            num nMoveType = 4
            num nPercentage
            num nSigValue = 1
        pointRx pPointRx[2]
        string sID
      [2]
        bool bMarked
        jointRx jJointRx = {j1=-87.551314, j2=145.129335, j3=-83.0857287, j4=182.11845, j5=63.691242, j6=-64.966659}
        pointRx pInter
        paraItem pParaItem
          [0]
            bool bSafePoint
            ifItem iIfItem
              [0]
                bool bANDOR[2]
                num nSigIndex[3]
                num nSigType[3]
                num nValue[3]
            mdesc mMdesc
            num nActionIndex = 42
            num nDelay
            num nMoveType = 1
            num nPercentage
            num nSigValue = 1
        pointRx pPointRx[2] = {x=61.349727, y=-652.129552, z=350.0734551, rx=-1.549449, ry=-1.96692, rz=28.421736, shoulder=lefty, elbow=enegative, wrist=wpositive}
        string sID
      [3]
        bool bMarked
        jointRx jJointRx = {j1=-47.00566362, j2=123.661152, j3=-79.978164, j4=176.739672, j5=50.379836, j6=-102.275032}
        pointRx pInter
        paraItem pParaItem
          [0]
            bool bSafePoint
            ifItem iIfItem
              [0]
                bool bANDOR[2]
                num nSigIndex[3]
                num nSigType[3]
                num nValue[3]
            mdesc mMdesc
            num nActionIndex = 42
            num nDelay
            num nMoveType = 1
            num nPercentage
            num nSigValue = 1
        pointRx pPointRx[2] = {x=488.627273, y=-418.649607, z=567.937104, rx=-6.582637, ry=-2.686226, rz=28.338446, shoulder=lefty, elbow=enegative, wrist=wpositive}
        string sID
      [4]
        bool bMarked
        jointRx jJointRx = {j1=-49.0942088, j2=121.00459063, j3=-74.169176, j4=177.183335, j5=53.609232, j6=-100.608132}
        pointRx pInter
        paraItem pParaItem
          [0]
            bool bSafePoint
            ifItem iIfItem
              [0]
                bool bANDOR[2]
                num nSigIndex[3]
                num nSigType[3]
                num nValue[3]
            mdesc mMdesc
            num nActionIndex = 42
            num nDelay
            num nMoveType = 1
            num nPercentage
            num nSigValue = 1
        pointRx pPointRx[2] = {x=488.602234, y=-457.380545, z=567.975681, rx=-6.584679, ry=-2.688341, rz=28.337484, shoulder=lefty, elbow=enegative, wrist=wpositive}
        string sID
      [5]
        bool bMarked
        jointRx jJointRx = {j1=-49.663191, j2=124.62488, j3=-82.121571, j4=177.0975297, j5=49.304971, j6=-99.821288}
        pointRx pInter
        paraItem pParaItem
          [0]
            bool bSafePoint
            ifItem iIfItem
              [0]
                bool bANDOR[2]
                num nSigIndex[3]
                num nSigType[3]
                num nValue[3]
            mdesc mMdesc
            num nActionIndex = 42
            num nDelay
            num nMoveType = 1
            num nPercentage
            num nSigValue = 1
        pointRx pPointRx[2] = {x=459.245528, y=-433.916408, z=567.993278, rx=-6.586651, ry=-2.689923, rz=28.337206, shoulder=lefty, elbow=enegative, wrist=wpositive}
        string sID
      [6]
        bool bMarked
        jointRx jJointRx = {j1=-51.089262, j2=127.485832, j3=-88.52739, j4=177.166583, j5=45.811078, j6=-98.322007}
        pointRx pInter
        paraItem pParaItem
          [0]
            bool bSafePoint
            ifItem iIfItem
              [0]
                bool bANDOR[2]
                num nSigIndex[3]
                num nSigType[3]
                num nValue[3]
            mdesc mMdesc
            num nActionIndex = 42
            num nDelay
            num nMoveType = 1
            num nPercentage
            num nSigValue = 1
        pointRx pPointRx[2] = {x=426.511567, y=-420.559077, z=567.993292, rx=-6.586458, ry=-2.69014, rz=28.337108, shoulder=lefty, elbow=enegative, wrist=wpositive}
        string sID
      [7]
        bool bMarked
        jointRx jJointRx = {j1=-53.0755743, j2=125.0272638, j3=-83.0148913, j4=177.619487, j5=48.919255, j6=-96.759929}
        pointRx pInter
        paraItem pParaItem
          [0]
            bool bSafePoint
            ifItem iIfItem
              [0]
                bool bANDOR[2]
                num nSigIndex[3]
                num nSigType[3]
                num nValue[3]
            mdesc mMdesc
            num nActionIndex = 42
            num nDelay
            num nMoveType = 1
            num nPercentage
            num nSigValue = 1
        pointRx pPointRx[2] = {x=426.51149, y=-458.270304, z=567.99328, rx=-6.585479, ry=-2.689619, rz=28.337033, shoulder=lefty, elbow=enegative, wrist=wpositive}
        string sID
      [8]
        bool bMarked
        jointRx jJointRx = {j1=-52.426636, j2=130.387774, j3=-95.172697, j4=177.208528, j5=42.11144, j6=-96.897847}
        pointRx pInter
        paraItem pParaItem
          [0]
            bool bSafePoint
            ifItem iIfItem
              [0]
                bool bANDOR[2]
                num nSigIndex[3]
                num nSigType[3]
                num nValue[3]
            mdesc mMdesc
            num nActionIndex = 42
            num nDelay
            num nMoveType = 1
            num nPercentage
            num nSigValue = 1
        pointRx pPointRx[2] = {x=393.481918, y=-402.66269, z=567.993281, rx=-6.585883, ry=-2.690348, rz=28.336908, shoulder=lefty, elbow=enegative, wrist=wpositive}
        string sID
      [9]
        bool bMarked
        jointRx jJointRx = {j1=-58.974439, j2=129.367388, j3=-92.816655, j4=178.435502, j5=43.592863, j6=-91.334255}
        pointRx pInter
        paraItem pParaItem
          [0]
            bool bSafePoint
            ifItem iIfItem
              [0]
                bool bANDOR[2]
                num nSigIndex[3]
                num nSigType[3]
                num nValue[3]
            mdesc mMdesc
            num nActionIndex = 42
            num nDelay
            num nMoveType = 1
            num nPercentage
            num nSigValue = 1
        pointRx pPointRx[2] = {x=344.945517, y=-458.235382, z=567.993294, rx=-6.587043, ry=-2.691097, rz=28.336907, shoulder=lefty, elbow=enegative, wrist=wpositive}
        string sID
      [10]
        bool bMarked
        jointRx jJointRx = {j1=-57.192018, j2=131.638959, j3=-98.096273, j4=178.00498558, j5=40.554749, j6=-92.720675}
        pointRx pInter
        paraItem pParaItem
          [0]
            bool bSafePoint
            ifItem iIfItem
              [0]
                bool bANDOR[2]
                num nSigIndex[3]
                num nSigType[3]
                num nValue[3]
            mdesc mMdesc
            num nActionIndex = 42
            num nDelay
            num nMoveType = 1
            num nPercentage
            num nSigValue = 1
        pointRx pPointRx[2] = {x=344.980685, y=-421.973821, z=567.993293, rx=-6.587471, ry=-2.690641, rz=28.337121, shoulder=lefty, elbow=enegative, wrist=wpositive}
        string sID
      [11]
        bool bMarked
        jointRx jJointRx = {j1=-60.376179, j2=132.512186, j3=-100.160991, j4=178.57184, j5=39.414626, j6=-89.972735}
        pointRx pInter
        paraItem pParaItem
          [0]
            bool bSafePoint
            ifItem iIfItem
              [0]
                bool bANDOR[2]
                num nSigIndex[3]
                num nSigType[3]
                num nValue[3]
            mdesc mMdesc
            num nActionIndex = 42
            num nDelay
            num nMoveType = 1
            num nPercentage
            num nSigValue = 1
        pointRx pPointRx[2] = {x=311.978155, y=-431.490165, z=567.993281, rx=-6.586244, ry=-2.690739, rz=28.336894, shoulder=lefty, elbow=enegative, wrist=wpositive}
        string sID
      [12]
        bool bMarked
        jointRx jJointRx = {j1=-65.107588, j2=132.458168, j3=-100.0326711, j4=179.493071, j5=39.531997, j6=-85.98983}
        pointRx pInter
        paraItem pParaItem
          [0]
            bool bSafePoint
            ifItem iIfItem
              [0]
                bool bANDOR[2]
                num nSigIndex[3]
                num nSigType[3]
                num nValue[3]
            mdesc mMdesc
            num nActionIndex = 42
            num nDelay
            num nMoveType = 1
            num nPercentage
            num nSigValue = 1
        pointRx pPointRx[2] = {x=270.822712, y=-458.161765, z=567.993281, rx=-6.586253, ry=-2.691371, rz=28.336679, shoulder=lefty, elbow=enegative, wrist=wpositive}
        string sID
      [13]
        bool bMarked
        jointRx jJointRx = {j1=-63.595033, j2=134.613161, j3=-105.229763, j4=179.141794, j5=36.481622, j6=-87.191501}
        pointRx pInter
        paraItem pParaItem
          [0]
            bool bSafePoint
            ifItem iIfItem
              [0]
                bool bANDOR[2]
                num nSigIndex[3]
                num nSigType[3]
                num nValue[3]
            mdesc mMdesc
            num nActionIndex = 42
            num nDelay
            num nMoveType = 1
            num nPercentage
            num nSigValue = 1
        pointRx pPointRx[2] = {x=270.822707, y=-423.00547317, z=567.99328, rx=-6.587117, ry=-2.691103, rz=28.336883, shoulder=lefty, elbow=enegative, wrist=wpositive}
        string sID
      [14]
        bool bMarked
        jointRx jJointRx = {j1=-65.403022, j2=136.841875, j3=-110.804443, j4=179.476622, j5=33.145897, j6=-85.649351}
        pointRx pInter
        paraItem pParaItem
          [0]
            bool bSafePoint
            ifItem iIfItem
              [0]
                bool bANDOR[2]
                num nSigIndex[3]
                num nSigType[3]
                num nValue[3]
            mdesc mMdesc
            num nActionIndex = 42
            num nDelay
            num nMoveType = 1
            num nPercentage
            num nSigValue = 1
        pointRx pPointRx[2] = {x=241.448098, y=-401.317138, z=567.99328, rx=-6.586652, ry=-2.691495, rz=28.336732, shoulder=lefty, elbow=enegative, wrist=wpositive}
        string sID
      [15]
        bool bMarked
        jointRx jJointRx = {j1=-71.552923, j2=137.207285, j3=-111.742738, j4=180.882707, j5=32.563572, j6=-80.728949}
        pointRx pInter
        paraItem pParaItem
          [0]
            bool bSafePoint
            ifItem iIfItem
              [0]
                bool bANDOR[2]
                num nSigIndex[3]
                num nSigType[3]
                num nValue[3]
            mdesc mMdesc
            num nActionIndex = 42
            num nDelay
            num nMoveType = 1
            num nPercentage
            num nSigValue = 1
        pointRx pPointRx[2] = {x=188.956768, y=-421.559208, z=567.993271, rx=-6.585305, ry=-2.691208, rz=28.336687, shoulder=lefty, elbow=enegative, wrist=wpositive}
        string sID
      [16]
        bool bMarked
        jointRx jJointRx = {j1=-72.731137, j2=135.0432437, j3=-106.287062, j4=181.0587207, j5=35.845376, j6=-79.673802}
        pointRx pInter
        paraItem pParaItem
          [0]
            bool bSafePoint
            ifItem iIfItem
              [0]
                bool bANDOR[2]
                num nSigIndex[3]
                num nSigType[3]
                num nValue[3]
            mdesc mMdesc
            num nActionIndex = 42
            num nDelay
            num nMoveType = 1
            num nPercentage
            num nSigValue = 1
        pointRx pPointRx[2] = {x=188.956768, y=-457.62638, z=567.99327, rx=-6.585271, ry=-2.690608, rz=28.336851, shoulder=lefty, elbow=enegative, wrist=wpositive}
        string sID
      [17]
        bool bMarked
        jointRx jJointRx = {j1=-75.0748224, j2=137.195165, j3=-111.715211, j4=181.688824, j5=32.546968, j6=-77.913471}
        pointRx pInter
        paraItem pParaItem
          [0]
            bool bSafePoint
            ifItem iIfItem
              [0]
                bool bANDOR[2]
                num nSigIndex[3]
                num nSigType[3]
                num nValue[3]
            mdesc mMdesc
            num nActionIndex = 42
            num nDelay
            num nMoveType = 1
            num nPercentage
            num nSigValue = 1
        pointRx pPointRx[2] = {x=159.184051, y=-433.850025, z=568.00311248, rx=-6.587391, ry=-2.691219, rz=28.336525, shoulder=lefty, elbow=enegative, wrist=wpositive}
        string sID
      [18]
        bool bMarked
        jointRx jJointRx = {j1=-79.693745, j2=136.402957, j3=-109.689565, j4=182.654161, j5=33.70043, j6=-74.112995}
        pointRx pInter
        paraItem pParaItem
          [0]
            bool bSafePoint
            ifItem iIfItem
              [0]
                bool bANDOR[2]
                num nSigIndex[3]
                num nSigType[3]
                num nValue[3]
            mdesc mMdesc
            num nActionIndex = 42
            num nDelay
            num nMoveType = 1
            num nPercentage
            num nSigValue = 1
        pointRx pPointRx[2] = {x=121.279103, y=-459.277382, z=568.00309762, rx=-6.585667, ry=-2.690876, rz=28.336551, shoulder=lefty, elbow=enegative, wrist=wpositive}
        string sID
      [19]
        bool bMarked
        jointRx jJointRx = {j1=-78.970374, j2=138.503231, j3=-115.146628, j4=182.739047, j5=30.363076, j6=-74.986334}
        pointRx pInter
        paraItem pParaItem
          [0]
            bool bSafePoint
            ifItem iIfItem
              [0]
                bool bANDOR[2]
                num nSigIndex[3]
                num nSigType[3]
                num nValue[3]
            mdesc mMdesc
            num nActionIndex = 42
            num nDelay
            num nMoveType = 1
            num nPercentage
            num nSigValue = 1
        pointRx pPointRx[2] = {x=121.279109, y=-423.991398, z=568.0031016, rx=-6.587075, ry=-2.690729, rz=28.336634, shoulder=lefty, elbow=enegative, wrist=wpositive}
        string sID
      [20]
        bool bMarked
        jointRx jJointRx = {j1=-82.18311, j2=140.325944, j3=-120.168865, j4=183.894102, j5=27.100815, j6=-72.899949}
        pointRx pInter
        paraItem pParaItem
          [0]
            bool bSafePoint
            ifItem iIfItem
              [0]
                bool bANDOR[2]
                num nSigIndex[3]
                num nSigType[3]
                num nValue[3]
            mdesc mMdesc
            num nActionIndex = 42
            num nDelay
            num nMoveType = 1
            num nPercentage
            num nSigValue = 1
        pointRx pPointRx[2] = {x=89.677736, y=-399.34141, z=568.00311271, rx=-6.587002, ry=-2.691537, rz=28.336424, shoulder=lefty, elbow=enegative, wrist=wpositive}
        string sID
      [21]
        bool bMarked
        jointRx jJointRx = {j1=-88.384098, j2=139.878985, j3=-118.905257, j4=185.387949, j5=27.7368, j6=-68.0421089}
        pointRx pInter
        paraItem pParaItem
          [0]
            bool bSafePoint
            ifItem iIfItem
              [0]
                bool bANDOR[2]
                num nSigIndex[3]
                num nSigType[3]
                num nValue[3]
            mdesc mMdesc
            num nActionIndex = 42
            num nDelay
            num nMoveType = 1
            num nPercentage
            num nSigValue = 1
        pointRx pPointRx[2] = {x=39.927338, y=-417.114199, z=568.00310299, rx=-6.585859, ry=-2.691076, rz=28.336552, shoulder=lefty, elbow=enegative, wrist=wpositive}
        string sID
      [22]
        bool bMarked
        jointRx jJointRx = {j1=-88.507848, j2=137.593086, j3=-112.746079, j4=184.812037, j5=31.590474, j6=-67.248671}
        pointRx pInter
        paraItem pParaItem
          [0]
            bool bSafePoint
            ifItem iIfItem
              [0]
                bool bANDOR[2]
                num nSigIndex[3]
                num nSigType[3]
                num nValue[3]
            mdesc mMdesc
            num nActionIndex = 42
            num nDelay
            num nMoveType = 1
            num nPercentage
            num nSigValue = 1
        pointRx pPointRx[2] = {x=39.927351, y=-456.440721, z=568.00310534, rx=-6.585835, ry=-2.690626, rz=28.33667, shoulder=lefty, elbow=enegative, wrist=wpositive}
        string sID
      [23]
        bool bMarked
        jointRx jJointRx = {j1=-92.775201, j2=139.648579, j3=-118.263421, j4=186.416179, j5=27.98427, j6=-64.573899}
        pointRx pInter
        paraItem pParaItem
          [0]
            bool bSafePoint
            ifItem iIfItem
              [0]
                bool bANDOR[2]
                num nSigIndex[3]
                num nSigType[3]
                num nValue[3]
            mdesc mMdesc
            num nActionIndex = 42
            num nDelay
            num nMoveType = 1
            num nPercentage
            num nSigValue = 1
        pointRx pPointRx[2] = {x=3.22242, y=-424.708167, z=568.00310073, rx=-6.587405, ry=-2.690621, rz=28.336622, shoulder=lefty, elbow=enegative, wrist=wpositive}
        string sID
      [24]
        bool bMarked
        jointRx jJointRx = {j1=-96.271776, j2=137.651223, j3=-112.897673, j4=186.564623, j5=31.174623, j6=-61.045352}
        pointRx pInter
        paraItem pParaItem
          [0]
            bool bSafePoint
            ifItem iIfItem
              [0]
                bool bANDOR[2]
                num nSigIndex[3]
                num nSigType[3]
                num nValue[3]
            mdesc mMdesc
            num nActionIndex = 42
            num nDelay
            num nMoveType = 1
            num nPercentage
            num nSigValue = 1
        pointRx pPointRx[2] = {x=-29.950899, y=-459.353258, z=568.00310491, rx=-6.585914, ry=-2.690721, rz=28.336673, shoulder=lefty, elbow=enegative, wrist=wpositive}
        string sID
      [25]
        bool bMarked
        jointRx jJointRx = {j1=-96.735861, j2=139.734616, j3=-118.502583, j4=187.433387, j5=27.658734, j6=-61.551893}
        pointRx pInter
        paraItem pParaItem
          [0]
            bool bSafePoint
            ifItem iIfItem
              [0]
                bool bANDOR[2]
                num nSigIndex[3]
                num nSigType[3]
                num nValue[3]
            mdesc mMdesc
            num nActionIndex = 42
            num nDelay
            num nMoveType = 1
            num nPercentage
            num nSigValue = 1
        pointRx pPointRx[2] = {x=-29.950895, y=-423.86666, z=568.00310038, rx=-6.587397, ry=-2.69039, rz=28.336676, shoulder=lefty, elbow=enegative, wrist=wpositive}
        string sID
      [26]
        bool bMarked
        jointRx jJointRx = {j1=-101.157848, j2=140.842973, j3=-121.666368, j4=189.150328, j5=25.409405, j6=-58.831913}
        pointRx pInter
        paraItem pParaItem
          [0]
            bool bSafePoint
            ifItem iIfItem
              [0]
                bool bANDOR[2]
                num nSigIndex[3]
                num nSigType[3]
                num nValue[3]
            mdesc mMdesc
            num nActionIndex = 42
            num nDelay
            num nMoveType = 1
            num nPercentage
            num nSigValue = 1
        pointRx pPointRx[2] = {x=-63.0350276, y=-401.658362, z=568.0119001, rx=-6.591358, ry=-2.690107, rz=28.336785, shoulder=lefty, elbow=enegative, wrist=wpositive}
        string sID
      [27]
        bool bMarked
        jointRx jJointRx = {j1=-106.321482, j2=139.390983, j3=-117.555756, j4=189.555383, j5=27.736636, j6=-53.876831}
        pointRx pInter
        paraItem pParaItem
          [0]
            bool bSafePoint
            ifItem iIfItem
              [0]
                bool bANDOR[2]
                num nSigIndex[3]
                num nSigType[3]
                num nValue[3]
            mdesc mMdesc
            num nActionIndex = 42
            num nDelay
            num nMoveType = 1
            num nPercentage
            num nSigValue = 1
        pointRx pPointRx[2] = {x=-111.697026, y=-421.905178, z=568.0118843, rx=-6.589731, ry=-2.690155, rz=28.336941, shoulder=lefty, elbow=enegative, wrist=wpositive}
        string sID
      [28]
        bool bMarked
        jointRx jJointRx = {j1=-105.163678, j2=137.182641, j3=-111.68623, j4=188.301748, j5=31.425495, j6=-53.655505}
        pointRx pInter
        paraItem pParaItem
          [0]
            bool bSafePoint
            ifItem iIfItem
              [0]
                bool bANDOR[2]
                num nSigIndex[3]
                num nSigType[3]
                num nValue[3]
            mdesc mMdesc
            num nActionIndex = 42
            num nDelay
            num nMoveType = 1
            num nPercentage
            num nSigValue = 1
        pointRx pPointRx[2] = {x=-111.697032, y=-459.394719, z=568.0118891, rx=-6.58976, ry=-2.689883, rz=28.337005, shoulder=lefty, elbow=enegative, wrist=wpositive}
        string sID
      [29]
        bool bMarked
        jointRx jJointRx = {j1=-109.993564, j2=138.161855, j3=-114.245931, j4=189.72279, j5=29.552893, j6=-50.212815}
        pointRx pInter
        paraItem pParaItem
          [0]
            bool bSafePoint
            ifItem iIfItem
              [0]
                bool bANDOR[2]
                num nSigIndex[3]
                num nSigType[3]
                num nValue[3]
            mdesc mMdesc
            num nActionIndex = 42
            num nDelay
            num nMoveType = 1
            num nPercentage
            num nSigValue = 1
        pointRx pPointRx[2] = {x=-149.400314, y=-435.0433995, z=568.0175242, rx=-6.593588, ry=-2.688525, rz=28.336857, shoulder=lefty, elbow=enegative, wrist=wpositive}
        string sID
      [30]
        bool bMarked
        jointRx jJointRx = {j1=-112.313327, j2=136.133118, j3=-109.0138371, j4=189.300283, j5=32.546465, j6=-47.276129}
        pointRx pInter
        paraItem pParaItem
          [0]
            bool bSafePoint
            ifItem iIfItem
              [0]
                bool bANDOR[2]
                num nSigIndex[3]
                num nSigType[3]
                num nValue[3]
            mdesc mMdesc
            num nActionIndex = 42
            num nDelay
            num nMoveType = 1
            num nPercentage
            num nSigValue = 1
        pointRx pPointRx[2] = {x=-181.55946, y=-459.58998, z=568.0175287, rx=-6.592761, ry=-2.688896, rz=28.33687, shoulder=lefty, elbow=enegative, wrist=wpositive}
        string sID
      [31]
        bool bMarked
        jointRx jJointRx = {j1=-113.964434, j2=138.396427, j3=-114.86875, j4=190.670185, j5=28.888812, j6=-47.13291}
        pointRx pInter
        paraItem pParaItem
          [0]
            bool bSafePoint
            ifItem iIfItem
              [0]
                bool bANDOR[2]
                num nSigIndex[3]
                num nSigType[3]
                num nValue[3]
            mdesc mMdesc
            num nActionIndex = 42
            num nDelay
            num nMoveType = 1
            num nPercentage
            num nSigValue = 1
        pointRx pPointRx[2] = {x=-181.594749, y=-421.537235, z=568.0175236, rx=-6.594319, ry=-2.688214, rz=28.336832, shoulder=lefty, elbow=enegative, wrist=wpositive}
        string sID
      [32]
        bool bMarked
        jointRx jJointRx = {j1=-118.604405, j2=138.501904, j3=-115.150042, j4=191.674761, j5=28.357416, j6=-43.427139}
        pointRx pInter
        paraItem pParaItem
          [0]
            bool bSafePoint
            ifItem iIfItem
              [0]
                bool bANDOR[2]
                num nSigIndex[3]
                num nSigType[3]
                num nValue[3]
            mdesc mMdesc
            num nActionIndex = 42
            num nDelay
            num nMoveType = 1
            num nPercentage
            num nSigValue = 1
        pointRx pPointRx[2] = {x=-218.976681, y=-405.617576, z=568.0175364, rx=-6.593482, ry=-2.689779, rz=28.336534, shoulder=lefty, elbow=enegative, wrist=wpositive}
        string sID
      [33]
        bool bMarked
        jointRx jJointRx = {j1=-122.43129, j2=136.510373, j3=-109.968352, j4=191.267208, j5=31.162627, j6=-38.960946}
        pointRx pInter
        paraItem pParaItem
          [0]
            bool bSafePoint
            ifItem iIfItem
              [0]
                bool bANDOR[2]
                num nSigIndex[3]
                num nSigType[3]
                num nValue[3]
            mdesc mMdesc
            num nActionIndex = 42
            num nDelay
            num nMoveType = 1
            num nPercentage
            num nSigValue = 1
        pointRx pPointRx[2] = {x=-266.781894, y=-418.843184, z=568.0175249, rx=-6.59271, ry=-2.689284, rz=28.336808, shoulder=lefty, elbow=enegative, wrist=wpositive}
        string sID
      [34]
        bool bMarked
        jointRx jJointRx = {j1=-120.363596, j2=134.220217, j3=-104.277478, j4=189.96233, j5=34.684647, j6=-39.577314}
        pointRx pInter
        paraItem pParaItem
          [0]
            bool bSafePoint
            ifItem iIfItem
              [0]
                bool bANDOR[2]
                num nSigIndex[3]
                num nSigType[3]
                num nValue[3]
            mdesc mMdesc
            num nActionIndex = 42
            num nDelay
            num nMoveType = 1
            num nPercentage
            num nSigValue = 1
        pointRx pPointRx[2] = {x=-266.781897, y=-456.916935, z=568.0175222, rx=-6.592282, ry=-2.68903, rz=28.336952, shoulder=lefty, elbow=enegative, wrist=wpositive}
        string sID
      [35]
        bool bMarked
        jointRx jJointRx = {j1=-125.0772856, j2=134.253942, j3=-104.360049, j4=190.690056, j5=34.21661, j6=-35.505136}
        pointRx pInter
        paraItem pParaItem
          [0]
            bool bSafePoint
            ifItem iIfItem
              [0]
                bool bANDOR[2]
                num nSigIndex[3]
                num nSigType[3]
                num nValue[3]
            mdesc mMdesc
            num nActionIndex = 42
            num nDelay
            num nMoveType = 1
            num nPercentage
            num nSigValue = 1
        pointRx pPointRx[2] = {x=-307.935358, y=-434.76833, z=568.017523, rx=-6.593883, ry=-2.688735, rz=28.336707, shoulder=lefty, elbow=enegative, wrist=wpositive}
        string sID
      [36]
        bool bMarked
        jointRx jJointRx = {j1=-126.18234, j2=131.562477, j3=-97.923448, j4=189.919943, j5=37.796067, j6=-33.392156}
        pointRx pInter
        paraItem pParaItem
          [0]
            bool bSafePoint
            ifItem iIfItem
              [0]
                bool bANDOR[2]
                num nSigIndex[3]
                num nSigType[3]
                num nValue[3]
            mdesc mMdesc
            num nActionIndex = 42
            num nDelay
            num nMoveType = 1
            num nPercentage
            num nSigValue = 1
        pointRx pPointRx[2] = {x=-339.344844, y=-459.232197, z=568.017529, rx=-6.592539, ry=-2.689542, rz=28.336769, shoulder=lefty, elbow=enegative, wrist=wpositive}
        string sID
      [37]
        bool bMarked
        jointRx jJointRx = {j1=-128.582305, j2=134.0504995, j3=-103.865016, j4=191.106968, j5=34.171376, j6=-32.340904}
        pointRx pInter
        paraItem pParaItem
          [0]
            bool bSafePoint
            ifItem iIfItem
              [0]
                bool bANDOR[2]
                num nSigIndex[3]
                num nSigType[3]
                num nValue[3]
            mdesc mMdesc
            num nActionIndex = 42
            num nDelay
            num nMoveType = 1
            num nPercentage
            num nSigValue = 1
        pointRx pPointRx[2] = {x=-339.309588, y=-418.740098, z=568.0175315, rx=-6.594008, ry=-2.688373, rz=28.336777, shoulder=lefty, elbow=enegative, wrist=wpositive}
        string sID
      [38]
        bool bMarked
        jointRx jJointRx = {j1=-132.557194, j2=133.634455, j3=-102.857498, j4=191.461094, j5=34.356586, j6=-28.624313}
        pointRx pInter
        paraItem pParaItem
          [0]
            bool bSafePoint
            ifItem iIfItem
              [0]
                bool bANDOR[2]
                num nSigIndex[3]
                num nSigType[3]
                num nValue[3]
            mdesc mMdesc
            num nActionIndex = 42
            num nDelay
            num nMoveType = 1
            num nPercentage
            num nSigValue = 1
        pointRx pPointRx[2] = {x=-375.559173, y=-400.058365, z=568.0175324, rx=-6.594143, ry=-2.688832, rz=28.336597, shoulder=lefty, elbow=enegative, wrist=wpositive}
        string sID
      [39]
        bool bMarked
        jointRx jJointRx = {j1=-119.478492, j2=120.691949, j3=-73.499146, j4=187.10756, j5=51.832735, j6=-36.651813}
        pointRx pInter
        paraItem pParaItem
          [0]
            bool bSafePoint
            ifItem iIfItem
              [0]
                bool bANDOR[2]
                num nSigIndex[3]
                num nSigType[3]
                num nValue[3]
            mdesc mMdesc
            num nActionIndex = 42
            num nDelay
            num nMoveType = 1
            num nPercentage
            num nSigValue = 1
        pointRx pPointRx[2] = {x=-337.807889, y=-600.36076, z=568.0175361, rx=-6.594662, ry=-2.688082, rz=28.336794, shoulder=lefty, elbow=enegative, wrist=wpositive}
        string sID
      [40]
        bool bMarked
        jointRx jJointRx = {j1=-114.66665, j2=123.31448, j3=-79.237868, j4=186.86886, j5=49.163146, j6=-41.566692}
        pointRx pInter
        paraItem pParaItem
          [0]
            bool bSafePoint
            ifItem iIfItem
              [0]
                bool bANDOR[2]
                num nSigIndex[3]
                num nSigType[3]
                num nValue[3]
            mdesc mMdesc
            num nActionIndex = 42
            num nDelay
            num nMoveType = 1
            num nPercentage
            num nSigValue = 1
        pointRx pPointRx[2] = {x=-270.459245, y=-600.323798, z=568.0421695, rx=-6.598641, ry=-2.685549, rz=28.337226, shoulder=lefty, elbow=enegative, wrist=wpositive}
        string sID
      [41]
        bool bMarked
        jointRx jJointRx = {j1=-107.974088, j2=125.672333, j3=-84.464513, j4=186.296074, j5=46.833882, j6=-48.0688486}
        pointRx pInter
        paraItem pParaItem
          [0]
            bool bSafePoint
            ifItem iIfItem
              [0]
                bool bANDOR[2]
                num nSigIndex[3]
                num nSigType[3]
                num nValue[3]
            mdesc mMdesc
            num nActionIndex = 42
            num nDelay
            num nMoveType = 1
            num nPercentage
            num nSigValue = 1
        pointRx pPointRx[2] = {x=-184.237317, y=-600.323785, z=568.0421684, rx=-6.598566, ry=-2.685446, rz=28.337311, shoulder=lefty, elbow=enegative, wrist=wpositive}
        string sID
      [42]
        bool bMarked
        jointRx jJointRx = {j1=-102.117608, j2=126.837266, j3=-87.076342, j4=185.596638, j5=45.789092, j6=-53.505467}
        pointRx pInter
        paraItem pParaItem
          [0]
            bool bSafePoint
            ifItem iIfItem
              [0]
                bool bANDOR[2]
                num nSigIndex[3]
                num nSigType[3]
                num nValue[3]
            mdesc mMdesc
            num nActionIndex = 42
            num nDelay
            num nMoveType = 1
            num nPercentage
            num nSigValue = 1
        pointRx pPointRx[2] = {x=-113.500018, y=-600.323774, z=568.0421674, rx=-6.598415, ry=-2.68541, rz=28.337367, shoulder=lefty, elbow=enegative, wrist=wpositive}
        string sID
      [43]
        bool bMarked
        jointRx jJointRx = {j1=-95.149611, j2=127.359728, j3=-88.254816, j4=184.578557, j5=45.528519, j6=-59.749811}
        pointRx pInter
        paraItem pParaItem
          [0]
            bool bSafePoint
            ifItem iIfItem
              [0]
                bool bANDOR[2]
                num nSigIndex[3]
                num nSigType[3]
                num nValue[3]
            mdesc mMdesc
            num nActionIndex = 42
            num nDelay
            num nMoveType = 1
            num nPercentage
            num nSigValue = 1
        pointRx pPointRx[2] = {x=-32.49609, y=-600.323763, z=568.0421666, rx=-6.598196, ry=-2.685321, rz=28.337443, shoulder=lefty, elbow=enegative, wrist=wpositive}
        string sID
      [44]
        bool bMarked
        jointRx jJointRx = {j1=-82.048942, j2=126.0420636, j3=-85.29102, j4=182.36613, j5=47.679346, j6=-71.157904}
        pointRx pInter
        paraItem pParaItem
          [0]
            bool bSafePoint
            ifItem iIfItem
              [0]
                bool bANDOR[2]
                num nSigIndex[3]
                num nSigType[3]
                num nValue[3]
            mdesc mMdesc
            num nActionIndex = 42
            num nDelay
            num nMoveType = 1
            num nPercentage
            num nSigValue = 1
        pointRx pPointRx[2] = {x=118.921487, y=-600.323741, z=568.0421643, rx=-6.597757, ry=-2.685415, rz=28.337426, shoulder=lefty, elbow=enegative, wrist=wpositive}
        string sID
      [45]
        bool bMarked
        jointRx jJointRx = {j1=-76.583274, j2=124.50583, j3=-81.872231, j4=181.422567, j5=49.681933, j6=-75.897744}
        pointRx pInter
        paraItem pParaItem
          [0]
            bool bSafePoint
            ifItem iIfItem
              [0]
                bool bANDOR[2]
                num nSigIndex[3]
                num nSigType[3]
                num nValue[3]
            mdesc mMdesc
            num nActionIndex = 42
            num nDelay
            num nMoveType = 1
            num nPercentage
            num nSigValue = 1
        pointRx pPointRx[2] = {x=184.871013, y=-600.305426, z=568.0561358, rx=-6.599219, ry=-2.684946, rz=28.351428, shoulder=lefty, elbow=enegative, wrist=wpositive}
        string sID
      [46]
        bool bMarked
        jointRx jJointRx = {j1=-64.919721, j2=118.302186, j3=-68.34286, j4=179.574591, j5=57.0732172, j6=-86.320686}
        pointRx pInter
        paraItem pParaItem
          [0]
            bool bSafePoint
            ifItem iIfItem
              [0]
                bool bANDOR[2]
                num nSigIndex[3]
                num nSigType[3]
                num nValue[3]
            mdesc mMdesc
            num nActionIndex = 42
            num nDelay
            num nMoveType = 1
            num nPercentage
            num nSigValue = 1
        pointRx pPointRx[2] = {x=339.597093, y=-600.305387, z=568.0561308, rx=-6.599008, ry=-2.684966, rz=28.351339, shoulder=lefty, elbow=enegative, wrist=wpositive}
        string sID
      [47]
        bool bMarked
        jointRx jJointRx = {j1=-55.452548, j2=107.0853304, j3=-44.666617, j4=178.376817, j5=69.385851, j6=-95.377402}
        pointRx pInter
        paraItem pParaItem
          [0]
            bool bSafePoint
            ifItem iIfItem
              [0]
                bool bANDOR[2]
                num nSigIndex[3]
                num nSigType[3]
                num nValue[3]
            mdesc mMdesc
            num nActionIndex = 42
            num nDelay
            num nMoveType = 1
            num nPercentage
